(* IEC 61131-3 sources: 2026_Projet_YGO_ExcavatriceDragage/CODE/E_CODEURS/_TYPES, 8 files *)

(* ---- E_PresetConfirmMode.st ---- *)
(* =======================================================================
   ⚙️ E_PresetConfirmMode — Mode de confirmation du preset codeur
   ───────────────────────────────────────────────────────────────────────
   🎯 Rôle : sélectionner le fait public utilisé pour valider un preset.
   📄 Doc : DOC/AF/AF_Partie-09_Fonction_Encoder_v2.4.md
   ======================================================================= *)

TYPE E_PresetConfirmMode :
ENUM
    READBACK_ONLY        := 0, // Confirmation par relecture de position
    READBACK_AND_STATUSBIT := 1, // Relecture et bit d'état matériel
    STATUSBIT_ONLY       := 2  // Bit d'état matériel uniquement
END_ENUM
END_TYPE

(* ---- ST_Encoder_Calib.st ---- *)
(* =======================================================================
   💾 ST_Encoder_Calib — Calibration & référence codeur (1 par treuil, RETAIN)
   ───────────────────────────────────────────────────────────────
   🎯 Rôle : Structure de calibration RETAIN par treuil (M1_EncoderCalib / M2_EncoderCalib)
   💾 Données : Références brutes, état homed et contrôle de cohérence redémarrage
   📄 Doc métier : DOC/AF/AF_Partie-09_Fonction_Encoder_v2.4.md
   ======================================================================= *)

TYPE ST_Encoder_Calib :
STRUCT
    // === DONNEES DE REFERENCE BRUTE (RETAIN) ===
    HomingRefRaw                 : UDINT;         // Valeur brute figee au dernier homing reussi
    LastKnownRawPos               : UDINT;         // Dernier point brut valide connu (continu)

    // === CONFIGURATION & REGLAGES TOLERANCE ===
    RestartCoherenceTolerancePts   : UDINT := 1000; // Tolerance redemarrage (pts, ~12% de 8192)

    // === ETATS DE CALIBRATION & SECURITE ===
    Homed                         : BOOL;          // TRUE des qu'un referencement a reussi
    HomingSuspect                 : BOOL;          // TRUE si incoherence detectee au redemarrage
    HomingProvisional             : BOOL;          // TRUE si zero provisoire 0m HX1 (avant HX4 8.5m)
END_STRUCT
END_TYPE

(* ---- ST_EncoderHw.st ---- *)
(* ═══════════════════════════════════════════════════════════════
   🔌 ST_EncoderHw — Frontière hardware codeur (IN/OUT)
   ───────────────────────────────────────────────────────────────
   🎯 Regroupe les entrées/sorties hardware d'un codeur absolu EtherCAT
      pour exposer l'interface physique de FB_Encoder de façon testable.
   🔌 Producteur/consommateur : PRG_02_Acquisition câble ce bus vers le device.
   📄 Doc : DOC/AF/AF_Partie-09_Fonction_Encoder_v2.4.md
   ═══════════════════════════════════════════════════════════════ *)
TYPE ST_EncoderHw :
STRUCT
    // === ENTREES BUS ETHERCAT (vers le codeur) ===
    RawPosIn            : UDINT;        // Position brute EtherCAT (in)
    AlarmsIn            : UINT;        // Codes alarmes bruts EtherCAT
    WarningsIn          : UINT;        // Codes avertissements bruts EtherCAT
    SlaveOperational    : BOOL;        // Esclave EtherCAT operationnel
    PresetAck           : BOOL;        // Pulse confirmation preset reussi
    PresetNak           : BOOL;        // Pulse echec / timeout preset

    // === SORTIES BUS (vers le codeur) ===
    PresetTriggerCmd    : WORD;        // Ordre declenchement preset vers PDO Rx
    CodeSeqTriggerCmd   : WORD;        // Ordre sequence code vers PDO Rx
    PresetValueOut      : UDINT;       // Valeur de preset transmise au PDO Rx
END_STRUCT
END_TYPE

(* ---- ST_EncoderMeasurements.st ---- *)
(* =======================================================================
   📊 ST_EncoderMeasurements — Mesures codeurs M1/M2 (contrat frontière)
   ───────────────────────────────────────────────────────────────
   ⚠️ ORPHELIN (Tâche C5 — nettoyage données mortes) : ce type n'est plus
   référencé par aucun consommateur dans le CODE actif (après consolidation
   bus acquisition I8, le bus ST_AcquisitionInterPrg utilise désormais
   EncoderM1/EncoderM2 : ST_AcquisitionEncoderQualified). CONSERVÉ (non
   supprimé) car référencé par le harnais de test TOOLS/TEST_AUTO_CI/
   registry.yaml (10 entrées) et par des artefacts bundle. → Proposé à
   l'archivage APRÈS mise à jour du harnais de test.
   ───────────────────────────────────────────────────────────────
   🎯 Rôle : Structure frontière regroupant les sous-DUTs de mesure des treuils M1 et M2
   🔌 Interface : Producteur unique PRG_02_Acquisition
   📄 Doc métier : DOC/AF/AF_Partie-06_Acquisition_Qualification_IO_v2.4.md
   ======================================================================= *)

TYPE ST_EncoderMeasurements :
STRUCT
    // === CHAINES DE MESURE PAR TREUIL ===
    M1 : ST_fbEncoder_Measurement; // Chaine de mesure treuil M1 (COD1)
    M2 : ST_fbEncoder_Measurement; // Chaine de mesure treuil M2 (COD2)
END_STRUCT
END_TYPE

(* ---- ST_fbEncoder_Cfg.st ---- *)
(* =======================================================================
   ⚙️ ST_fbEncoder_Cfg — Réglages technologiques publics de FB_Encoder
   ───────────────────────────────────────────────────────────────────────
   🎯 Rôle : porter le mode de confirmation preset commun aux codeurs.
   🔒 Ownership : GVL_IHM.Commun.EncoderCfg ↔ GVL_PERSISTENT._EncoderCfgPersist.
   📄 Doc : DOC/AF/AF_Partie-09_Fonction_Encoder_v2.4.md
   ======================================================================= *)

TYPE ST_fbEncoder_Cfg :
STRUCT
    PresetConfirmMode : E_PresetConfirmMode := E_PresetConfirmMode.READBACK_ONLY; // Mode de confirmation preset, défaut relecture
    Initialized       : BOOL := FALSE;                        // 🚦 TRUE après restauration du pont persistant
END_STRUCT
END_TYPE

(* ---- ST_fbEncoder_HwIn.st ---- *)
(* =======================================================================
   🔌 ST_fbEncoder_HwIn — Faits hardware d'entrée codeur (HwIn)
   ───────────────────────────────────────────────────────────────
   🎯 Rôle : Regrouper les SEULES entrées/faits hardware d'un codeur absolu
      EtherCAT consommés par FB_Encoder (lecture seule côté automate).
   🔒 Ownership : PRG_02_Acquisition câble ce bus depuis le device/simulé.
   🛡️ PresetStatusBit : bit du mot d'état codeur, réservé site futur —
      câblé à FALSE tant qu'aucun bit n'est identifié (aucun signal absent
      ne confirme implicitement le preset).
   📄 Doc métier : DOC/AF/AF_Partie-09_Fonction_Encoder_v2.4.md
   ======================================================================= *)

TYPE ST_fbEncoder_HwIn :
STRUCT
    // === ENTRÉES BUS ETHERCAT (faits d'entrée, lecture seule) ===
    RawPosIn           : UDINT; // --> [HW] Position brute codeur
    SpdValueIn         : DINT;  // --> [HW] Vitesse brute codeur (0x6031:01 en 0.1 RPM)
    AlarmsIn           : UINT;  // --> [HW] Alarmes brutes codeur
    WarningsIn         : UINT;  // --> [HW] Avertissements bruts codeur
    SlaveOperational   : BOOL;  // --> [HW] Esclave EtherCAT operationnel
    PresetStatusBit    : BOOL;  // --> [HW] Bit d'etat preset optionnel, FALSE si non cable
END_STRUCT
END_TYPE

(* ---- ST_fbEncoder_HwOut.st ---- *)
(* =======================================================================
   🔌 ST_fbEncoder_HwOut — Ordres preset de sortie codeur (HwOut)
   ───────────────────────────────────────────────────────────────
   🎯 Rôle : Regrouper les SEULES sorties/ordres preset d'un codeur absolu
      EtherCAT produits par FB_Encoder vers le PDO Rx (bus sortie).
   🔒 Ownership : FB_Encoder produit ce bus ; PRG_02_Acquisition le relaie
      vers le device.
   📄 Doc métier : DOC/AF/AF_Partie-09_Fonction_Encoder_v2.4.md
   ======================================================================= *)

TYPE ST_fbEncoder_HwOut :
STRUCT
    // === SORTIES BUS ETHERCAT (ordres preset vers PDO Rx) ===
    PresetTriggerCmd   : WORD;   // <-- [ACT] Declenchement preset vers PDO Rx
    CodeSeqTriggerCmd  : WORD;   // <-- [ACT] Sequence code vers PDO Rx, maintenue a 0
    PresetValueOut     : UDINT;  // <-- [ACT] Valeur brute envoyee au preset
END_STRUCT
END_TYPE

(* ---- ST_fbEncoder_Measurement.st ---- *)
(* =======================================================================
   📊 ST_fbEncoder_Measurement — Mesures codeur conditionnées (1 sous-DUT par treuil)
   ───────────────────────────────────────────────────────────────
   🎯 Rôle : Regroupement des mesures et faits de la chaîne codeur d'un treuil (Abs → Scale → Safety → Speed)
   🔌 Interface : Interface de mesure normalisée pour PRG_02_Acquisition
   📄 Doc métier : DOC/AF/AF_Partie-06_Acquisition_Qualification_IO_v2.4.md
   ======================================================================= *)

TYPE ST_fbEncoder_Measurement :
STRUCT
    // === DONNEES BRUTES & STATUT BUS ===
    RawPos            : UDINT;        // Position brute codeur (gelee si EncoderAvailable=FALSE)
    EncoderAvailable  : BOOL;         // TRUE = bus/esclave EtherCAT operationnel et disponible

    // === MESURES DE POSITION CABLE ===
    CablePosM         : REAL;         // Position cable (m, signee, + enroule)
    CablePosMSafe     : REAL;         // Position cable instantanee validee par EncoderIncoherent (m)
    EncoderIncoherent : BOOL;         // TRUE = incoherence redemarrage ou hors bornes

    // === MESURES DE VITESSE CABLE ===
    Speed_Mps         : REAL;         // Vitesse absolue câble (m/s)
    SignedSpeed_Mps   : REAL;         // Vitesse signee câble (m/s, + montee, - descente)
    SpeedValid        : BOOL;         // TRUE si mesure valide et codeur operationnel

    // === STATUTS DES SOUS-FB & REFERENCE ===
    HomingFault       : ST_Fault;     // Défaut FB_Encoder_Homing (état du référencement)
    HomingLifecycle   : ST_Lifecycle; // Cycle FB_Encoder_Homing (Busy/Done)
    AbsFault          : ST_Fault;     // Défaut FB_Encoder_Abs (état acquisition bus)
    HomingRefRaw      : UDINT;        // Reference brute du dernier homing reussi (re-expose)
END_STRUCT
END_TYPE
